Fanuc KAREL source: ka00165.KL

-- PROVISIONAL review KL for V940-1; original PC SHA256 3319d7f71ef8fcdd9baad7429b3cda2eba6fc9e94638ff0f8c58afd57ffe4d83
-- Incomplete behavior may be omitted. Consult companion uncertainty JSON. Do not deploy.
PROGRAM KA00165
%NOLOCKGROUP
-- UNRESOLVED_DECL SRC type=002012
-- UNRESOLVED_DECL DST type=002012
BEGIN
  -- V9_COMPOSED_GLOBAL_TRANSFER_HINT repetitions=1; address IDs observed; pairing/direction/source/runtime held
  -- V9_TWO_GLOBAL_ADDRESS_COPY_HINT bounded five-record physical form; type/direction/source/runtime held
  -- V9_ZERO_TABLE_METADATA_HINT layout=0001; no indexed target words; source/name/runtime held
  -- UNRESOLVED_PC offsets 5-19; opcodes 22,22,1E
  -- UNRESOLVED_PC offsets 24-28; opcodes 7F
END KA00165
